{attribute 'enable_dynamic_creation'}
FUNCTION_BLOCK FB_TraceId IMPLEMENTS I_OtlpValue
VAR_OUTPUT
	bytes: ARRAY [0..15] OF BYTE;
END_VAR

(*
	Releases this value and clears the caller's pointer to it: call it as p^.delete(pSelf:=p).
	pSelf is cleared before the value is freed, so the caller never keeps a dangling pointer.
	A pointer to any other object is refused and left untouched, and nothing is released.
*)
METHOD delete : BOOL
VAR_IN_OUT
	pSelf: POINTER TO FB_TraceId;
END_VAR
VAR
	_pThis: POINTER TO FB_TraceId;
END_VAR
_pThis := THIS;
IF pSelf <> _pThis THEN
	RETURN;
END_IF

pSelf := 0;
__DELETE(_pThis);
delete := TRUE;
END_METHOD

PROPERTY eType : E_ValueType
GET
eType := E_ValueType.E_TraceId;
END_GET
END_PROPERTY

//FB_Exit must be implemented explicitly. If there is an implementation, then the
//method is called before the controller removes the code of the function block instance
//(implicit call). The return value is not evaluated.
METHOD FB_Exit: BOOL
VAR_INPUT
    bInCopyCode: BOOL;  // TRUE: the exit method is called in order to leave the instance which will be copied afterwards (online change).  
END_VAR
THIS^.free();
END_METHOD

METHOD free
// just resets values to defaults
MEMSET(ADR(THIS^.bytes), 0, SIZEOF(THIS^.bytes));
END_METHOD

END_FUNCTION_BLOCK

(* stored: Version 1.1.0.1
   POU FB_TraceId: Id {957763e9-1dc3-43f7-8bee-d4f8556d5952}, SpecialFunc None
   Method delete: Id {c97e0256-4d82-467f-8451-1a78cc35cf61}
   Property eType: Id {a8e38517-e28e-4988-8201-c1e2d19bf319}
   Get Get: Id {932f2685-55a3-403d-b638-288e54b28a9f}
   Method FB_Exit: Id {c97eaf69-2ccb-4370-a9b2-610f66a40aba}
   Method free: Id {f2521e9b-00ca-4214-9c98-a50a3ee6d37e} *)
